// TIA Portal V21 export
Screen "R09_Bar"  1024x768, Number=49, Template=Tpl
  ScreenLayer 
    Bar "P_Bar" at 10,10 size 100x30  MaximumValue=24
      ProcessValue := P_Cell
